// TIA Portal V20 export
Screen "Pop-up_TEC_UNIT_LEGEND_Popup"  400x487
  ScreenItem "Background" at 0,0 size 400x487  Type=HmiRectangle
  ScreenItem "Textfeld_Legende" at 1,1 size 398x25  Type=HmiTextBox
  ScreenItem "Arrow_ADV_Left_Fast" at 10,207 size 15x30  Type=HmiPolygon
  ScreenItem "Arrow_RTN_Right_Fast" at 40,207 size 15x30  Type=HmiPolygon
  ScreenItem "Arrow_RTN_Up_Fast" at 10,256 size 30x15  Type=HmiPolygon
  ScreenItem "Arrow_ADV_Down_Fast" at 40,256 size 30x15  Type=HmiPolygon
  ScreenItem "Textfeld_2" at 10,138 size 165x20  Type=HmiTextBox
  ScreenItem "Textfeld_1" at 10,160 size 165x20  Type=HmiTextBox
  ScreenItem "Textfeld_3" at 10,33 size 165x20  Type=HmiTextBox
  ScreenItem "Textfeld_4" at 10,55 size 165x20  Type=HmiTextBox
  ScreenItem "Textfeld_5" at 10,85 size 165x20  Type=HmiTextBox
  ScreenItem "Textfeld_6" at 10,117 size 165x20  Type=HmiTextBox
  ScreenItem "Rechteck_2" at 10,292 size 20x20  Type=HmiRectangle
  ScreenItem "Rechteck_5" at 10,328 size 40x10  Type=HmiRectangle
  ScreenItem "Grafikanzeige_1" at 10,371 size 16x16  Type=HmiGraphicView
  ScreenItem "Textfeld_7" at 10,412 size 20x20  Type=HmiTextBox
  ScreenItem "Textfeld_8" at 10,452 size 20x20  Type=HmiTextBox
  ScreenItem "Textfeld_9" at 180,138 size 165x20  Type=HmiTextBox
  ScreenItem "Textfeld_10" at 180,160 size 165x20  Type=HmiTextBox
  ScreenItem "Textfeld_11" at 180,33 size 117x20  Type=HmiTextBox
  ScreenItem "Textfeld_12" at 180,55 size 120x20  Type=HmiTextBox
  ScreenItem "Textfeld_13" at 180,77 size 215x37  Type=HmiTextBox
  ScreenItem "Textfeld_14" at 180,117 size 165x20  Type=HmiTextBox
  ScreenItem "Textfeld_15" at 10,185 size 100x20  Type=HmiTextBox
  ScreenItem "Textfeld_16" at 75,204 size 315x37  Type=HmiTextBox
  ScreenItem "Textfeld_17" at 75,244 size 315x40  Type=HmiTextBox
  ScreenItem "Textfeld_18" at 75,283 size 315x37  Type=HmiTextBox
  ScreenItem "Textfeld_19" at 75,324 size 315x37  Type=HmiTextBox
  ScreenItem "Textfeld_20" at 75,363 size 315x37  Type=HmiTextBox
  ScreenItem "Textfeld_21" at 75,403 size 315x37  Type=HmiTextBox
  ScreenItem "Textfeld_22" at 75,443 size 315x37  Type=HmiTextBox
  ScreenItem "Cancel Mode" at 309,1 size 90x60  Type=HmiButton
  ScreenItem "Rechteck_3" at 40,292 size 20x20  Type=HmiRectangle
  ScreenItem "Rechteck_4" at 10,348 size 40x10  Type=HmiRectangle
  ScreenItem "Textfeld_23" at 40,412 size 20x20  Type=HmiTextBox
  ScreenItem "Textfeld_24" at 40,452 size 20x20  Type=HmiTextBox
